(* IEC 61131-3 sources: HydroSim/openplc, 7 files *)

(* ---- watertanklogica.st ---- *)
PROGRAM program0
  VAR
    LowLevelSensor AT %IX0.5 : BOOL;
    ZoneAButton AT %IX0.6 : BOOL;
    ZoneBButton AT %IX0.7 : BOOL;
    ZoneCButton AT %IX1.0 : BOOL;
    ZoneDButton AT %IX1.1 : BOOL;
    HighLevelSensor AT %IX0.4 : BOOL;
    OverFlowSensor AT %IX0.3 : BOOL;
    Pump AT %QX0.1 : BOOL;
    Alarm AT %QX0.0 : BOOL;
    StartButton AT %IX0.0 : BOOL;
    StopButton AT %IX0.1 : BOOL;
    DrainButton AT %IX0.2 : BOOL;
    DrainValve AT %QX0.3 : BOOL;
    ValveZoneA AT %QX0.4 : BOOL;
    ValveZoneB AT %QX0.5 : BOOL;
    ValveZoneC AT %QX0.6 : BOOL;
    ValveZoneD AT %QX0.7 : BOOL;
  END_VAR

  Pump := NOT(StopButton) AND (Pump OR (LowLevelSensor AND StartButton));
  Alarm := OverFlowSensor;
  DrainValve := DrainButton AND NOT(LowLevelSensor);
  ValveZoneA := ZoneAButton;
  ValveZoneB := ZoneBButton;
  ValveZoneC := ZoneCButton;
  ValveZoneD := ZoneDButton;
END_PROGRAM

CONFIGURATION Config0

  RESOURCE Res0 ON PLC
    TASK task0(INTERVAL := T#20ms, PRIORITY := 0);
    PROGRAM instance0 WITH task0 : program0;
  END_RESOURCE
END_CONFIGURATION

(* ---- waterwijklogica.st ---- *)
PROGRAM program0
  VAR
    StartSwitch AT %IX0.0 : BOOL := TRUE;
    LowPressureSensor AT %IX0.1 : BOOL;
    HighPressureSensor AT %IX0.2 : BOOL;
    FaultSensor AT %IX0.3 : BOOL;
    EmergencyStop AT %IX0.4 : BOOL;
    MainPump AT %QX0.0 : BOOL;
    Alarm AT %QX0.1 : BOOL;
    PumpSpeed AT %MD1000 : REAL;
    PumpSpeedBits AT %MD1006 : DWORD;
    Pump1SpeedHigh AT %QW1000 : WORD;
    Pump1SpeedLow AT %QW1001 : WORD;
    Pump2SpeedHigh AT %QW1002 : WORD;
    Pump2SpeedLow AT %QW1003 : WORD;
    Pump3SpeedHigh AT %QW1004 : WORD;
    Pump3SpeedLow AT %QW1005 : WORD;
  END_VAR

  MainPump := StartSwitch;
  Alarm := FaultSensor OR EmergencyStop;

  IF MainPump THEN
    PumpSpeed := 1.0;
  ELSE
    PumpSpeed := 0.0;
  END_IF;

  PumpSpeedBits := REAL_TO_DWORD(PumpSpeed);
  Pump1SpeedHigh := DWORD_TO_WORD(SHR(IN := PumpSpeedBits, N := 16));
  Pump1SpeedLow := DWORD_TO_WORD(PumpSpeedBits AND DWORD#16#0000FFFF);
  Pump2SpeedHigh := Pump1SpeedHigh;
  Pump2SpeedLow := Pump1SpeedLow;
  Pump3SpeedHigh := Pump1SpeedHigh;
  Pump3SpeedLow := Pump1SpeedLow;
END_PROGRAM

CONFIGURATION Config0

  RESOURCE Res0 ON PLC
    TASK task0(INTERVAL := T#20ms, PRIORITY := 0);
    PROGRAM instance0 WITH task0 : program0;
  END_RESOURCE
END_CONFIGURATION

(* ---- zone_0.st ---- *)
PROGRAM Zone0Logica
  VAR
    Pump0_Run AT %QX0.0 : BOOL;
    Pump1_Run AT %QX0.1 : BOOL;
    Pump2_Run AT %QX0.2 : BOOL;
    Pump3_Run AT %QX0.3 : BOOL;

    Pump0_Cmd AT %QX0.4 : BOOL;
    Pump1_Cmd AT %QX0.5 : BOOL;
    Pump2_Cmd AT %QX0.6 : BOOL;
    Pump3_Cmd AT %QX0.7 : BOOL;

    Valve0_Run AT %QX1.0 : BOOL;
    Valve1_Run AT %QX1.1 : BOOL;
    Valve2_Run AT %QX1.2 : BOOL;
    Valve3_Run AT %QX1.3 : BOOL;
    Valve4_Run AT %QX1.4 : BOOL;
    Valve5_Run AT %QX1.5 : BOOL;
    Valve6_Run AT %QX1.6 : BOOL;
    Valve7_Run AT %QX1.7 : BOOL;
    Valve8_Run AT %QX2.0 : BOOL;

    Valve0_Cmd AT %QX2.1 : BOOL;
    Valve1_Cmd AT %QX2.2 : BOOL;
    Valve2_Cmd AT %QX2.3 : BOOL;
    Valve3_Cmd AT %QX2.4 : BOOL;
    Valve4_Cmd AT %QX2.5 : BOOL;
    Valve5_Cmd AT %QX2.6 : BOOL;
    Valve6_Cmd AT %QX2.7 : BOOL;
    Valve7_Cmd AT %QX3.0 : BOOL;
    Valve8_Cmd AT %QX3.1 : BOOL;

    T0_Low AT %IX0.0 : BOOL;
    T0_High AT %IX0.1 : BOOL;

    T1_High AT %IX0.2 : BOOL;
    T1_Low AT %IX0.3 : BOOL;

    T2_High AT %IX0.4 : BOOL;
    T2_Low AT %IX0.5 : BOOL;

    T3_High AT %IX0.6 : BOOL;
    T3_Low AT %IX0.7 : BOOL;

  END_VAR

  Valve0_Run := Valve0_Cmd;
  Valve1_Run := Valve1_Cmd;
  Valve2_Run := Valve2_Cmd;
  Valve3_Run := Valve3_Cmd;
  Valve4_Run := Valve4_Cmd;
  Valve5_Run := Valve5_Cmd;
  Valve6_Run := Valve6_Cmd;
  Valve7_Run := Valve7_Cmd;
  Valve8_Run := Valve8_Cmd;
  IF Valve0_Run = 0 THEN
    Pump0_Cmd := 0;
    Pump1_Cmd := 0;
    Pump2_Cmd := 0;
    Pump3_Cmd := 0;
  END_IF;

  Pump0_Run := Pump0_Cmd;
  Pump1_Run := Pump1_Cmd;
  Pump2_Run := Pump2_Cmd;
  Pump3_Run := Pump3_Cmd;
END_PROGRAM

CONFIGURATION Config0
  RESOURCE Res0 ON PLC
    TASK TaskMain(INTERVAL := T#50ms,PRIORITY := 0);
    PROGRAM Inst0 WITH TaskMain : Zone0Logica;
  END_RESOURCE
END_CONFIGURATION

(* ---- zone_1.st ---- *)
PROGRAM Zone1Logica
  VAR
    Pump_Run AT %QX0.0 : BOOL;
    Pump_Cmd AT %QX0.1 : BOOL;

    Valve0_Run AT %QX0.2 : BOOL;
    Valve0_Cmd AT %QX0.3 : BOOL;

    Valve1_Run AT %QX0.4 : BOOL;
    Valve1_Cmd AT %QX0.5 : BOOL;
  END_VAR

  Pump_Run := Pump_Cmd;
  Valve0_Run := Valve0_Cmd;
  Valve1_Run := Valve1_Cmd;

  IF Valve0_Run = FALSE THEN
    Pump_Cmd := FALSE;
  END_IF;
END_PROGRAM

CONFIGURATION Config0
  RESOURCE Res0 ON PLC
    TASK TaskMain(INTERVAL := T#50ms,PRIORITY := 0);
    PROGRAM Inst0 WITH TaskMain : Zone1Logica;
  END_RESOURCE
END_CONFIGURATION

(* ---- zone_2.st ---- *)
PROGRAM Zone2Logica
  VAR
    Pump_Run AT %QX0.0 : BOOL;
    Pump_Cmd AT %QX0.1 : BOOL;

    Valve0_Run AT %QX0.2 : BOOL;
    Valve0_Cmd AT %QX0.3 : BOOL;

    Valve1_Run AT %QX0.4 : BOOL;
    Valve1_Cmd AT %QX0.5 : BOOL;
  END_VAR

  Pump_Run := Pump_Cmd;
  Valve0_Run := Valve0_Cmd;
  Valve1_Run := Valve1_Cmd;

  IF Valve0_Run = FALSE THEN
    Pump_Cmd := FALSE;
  END_IF;
END_PROGRAM

CONFIGURATION Config0
  RESOURCE Res0 ON PLC
    TASK TaskMain(INTERVAL := T#50ms,PRIORITY := 0);
    PROGRAM Inst0 WITH TaskMain : Zone2Logica;
  END_RESOURCE
END_CONFIGURATION

(* ---- zone_3.st ---- *)
PROGRAM Zone3Logica
  VAR
    Pump_Run AT %QX0.0 : BOOL;
    Pump_Cmd AT %QX0.1 : BOOL;

    Valve0_Run AT %QX0.2 : BOOL;
    Valve0_Cmd AT %QX0.3 : BOOL;

    Valve1_Run AT %QX0.4 : BOOL;
    Valve1_Cmd AT %QX0.5 : BOOL;
  END_VAR

  Pump_Run := Pump_Cmd;
  Valve0_Run := Valve0_Cmd;
  Valve1_Run := Valve1_Cmd;

  IF Valve0_Run = FALSE THEN
    Pump_Cmd := FALSE;
  END_IF;
END_PROGRAM

CONFIGURATION Config0
  RESOURCE Res0 ON PLC
    TASK TaskMain(INTERVAL := T#50ms,PRIORITY := 0);
    PROGRAM Inst0 WITH TaskMain : Zone3Logica;
  END_RESOURCE
END_CONFIGURATION

(* ---- zone_4.st ---- *)
PROGRAM Zone4Logica
  VAR
    Pump_Run AT %QX0.0 : BOOL;
    Pump_Cmd AT %QX0.1 : BOOL;

    Valve0_Run AT %QX0.2 : BOOL;
    Valve0_Cmd AT %QX0.3 : BOOL;

    Valve1_Run AT %QX0.4 : BOOL;
    Valve1_Cmd AT %QX0.5 : BOOL;
  END_VAR

  Pump_Run := Pump_Cmd;
  Valve0_Run := Valve0_Cmd;
  Valve1_Run := Valve1_Cmd;

  IF Valve0_Run = FALSE THEN
    Pump_Cmd := FALSE;
  END_IF;
END_PROGRAM

CONFIGURATION Config0
  RESOURCE Res0 ON PLC
    TASK TaskMain(INTERVAL := T#50ms,PRIORITY := 0);
    PROGRAM Inst0 WITH TaskMain : Zone4Logica;
  END_RESOURCE
END_CONFIGURATION
